NAMESPACE TiaMcp_UnitA
DATA_BLOCK "TgpUnit_GlobalTimer"
{ S7_Optimized_Access := 'TRUE' }
VERSION : 0.1
"IEC_TIMER"
BEGIN
END_DATA_BLOCK

DATA_BLOCK "TgpUnit_GlobalCounter"
{ S7_Optimized_Access := 'TRUE' }
VERSION : 0.1
"IEC_COUNTER"
BEGIN
END_DATA_BLOCK

DATA_BLOCK "TgpUnit_NumericFB_DB"
{ S7_Optimized_Access := 'TRUE' }
VERSION : 0.1
"TgpUnit_NumericFB"
BEGIN
END_DATA_BLOCK

DATA_BLOCK "TgpUnit_GlobalTemplateFB_LAD"
{ S7_Optimized_Access := 'TRUE' }
VERSION : 0.1
"TgpUnit_TemplateFB_LAD"
BEGIN
END_DATA_BLOCK

DATA_BLOCK "TgpUnit_GlobalTemplateFB_FBD"
{ S7_Optimized_Access := 'TRUE' }
VERSION : 0.1
"TgpUnit_TemplateFB_FBD"
BEGIN
END_DATA_BLOCK

FUNCTION_BLOCK "TgpUnit_MultiTemplateFB_LAD"
{ S7_Optimized_Access := 'TRUE' }
VERSION : 0.1
VAR
 Child : "TgpUnit_TemplateFB_LAD";
END_VAR
BEGIN
END_FUNCTION_BLOCK

FUNCTION_BLOCK "TgpUnit_MultiTemplateFB_FBD"
{ S7_Optimized_Access := 'TRUE' }
VERSION : 0.1
VAR
 Child : "TgpUnit_TemplateFB_FBD";
END_VAR
BEGIN
END_FUNCTION_BLOCK

END_NAMESPACE
